(*
    States of FB_FemtoAmplifier, reported as Status.State (code) and
    Status.StateText (name).
*)
{attribute 'qualified_only'}
{attribute 'strict'}
{attribute 'to_string'}
TYPE E_FemtoState :
(
    READY := 0,     // settings in use have settled
    SETTLING := 1   // within the settling time after a change or a PLC start
);
END_TYPE

(* stored: Version 1.1.0.1
   DUT E_FemtoState: Id {f04d0066-4206-4a9e-8cbb-a17a967434b3} *)
